ADAPTER pos_init (* Adapter Interface *)
  (* Standard: 61499-1 *)
  (* Version 0.0, 10/22/2026, macie, Schneider Electric *)
  PACKAGE Main;
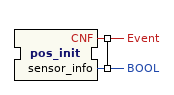
  EVENT_OUTPUT
    CNF WITH sensor_info; (* Confirmation from Plug *)
  END_EVENT
  VAR_OUTPUT
    sensor_info : BOOL; (* Confirmation Data from Plug *)
  END_VAR
  SERVICE SOCKET/PLUG
    SEQUENCE request_confirm
      SOCKET.REQ(REQD) -> PLUG.REQ(REQD);
      PLUG.CNF(sensor_info) -> SOCKET.CNF(sensor_info);
    END_SEQUENCE
    SEQUENCE indication_response
      PLUG.IND(INDD) -> SOCKET.IND(INDD);
      SOCKET.RSP(RSPD) -> PLUG.RSP(RSPD);
    END_SEQUENCE
  END_SERVICE
END_ADAPTER
